Fanuc KAREL source: kt00604.KL

-- PROVISIONAL review KL for V770-1; original PC SHA256 ef8bddbbafa6d18c365e844a8c896fe21d5d31c39a11a245256090b743b57c69
-- Incomplete behavior may be omitted. Consult companion uncertainty JSON. Do not deploy.
PROGRAM KT00604
%NOLOCKGROUP
VAR
  I1 : INTEGER
  I2 : INTEGER
  OUT : INTEGER
BEGIN
  -- UNRESOLVED_PC offsets 5-16; opcodes 2E,23
  -- UNRESOLVED_PC offsets 21-32; opcodes 2E,23
  -- UNRESOLVED_PC offsets 37-48; opcodes 2E,23
  -- UNRESOLVED_PC offsets 53-64; opcodes 2E,23
  -- UNRESOLVED_PC offsets 69-82; opcodes 21,51,23
  -- UNRESOLVED_PC offsets 87-91; opcodes 7F
END KT00604
